(* IEC 61131-3 sources: plc-iiot-stack/tests/POUs/F_TestContains, 2 files *)

(* ---- F_TestContains.decl.st ---- *)
// Назначение: для тестов — содержит ли текст длиной до MQTT_PAYLOAD_LEN подстроку sPart (стандартная
//             FIND работает только со строками до 255 символов).
// Автор:      kr0nsch
// Версия:     0.1.0
// Документ:   docs/TEST_REPORT.md
FUNCTION F_TestContains : BOOL
VAR_IN_OUT CONSTANT
    // lint:allow STL007 параметр VAR_IN_OUT CONSTANT — ссылка только для чтения, а не константа
    sText : STRING(GVL_Const.MQTT_PAYLOAD_LEN);
END_VAR
VAR_INPUT
    sPart : STRING(255);
END_VAR
VAR
    uiTextLen : UINT;
    uiPartLen : UINT;
    uiStart : UINT;
    uiIdx : UINT;
    xMatch : BOOL;
END_VAR

(* ---- F_TestContains.impl.st ---- *)
uiPartLen := INT_TO_UINT(LEN(sPart));
uiTextLen := 0;
WHILE uiTextLen < GVL_Const.MQTT_PAYLOAD_LEN AND_THEN sText[uiTextLen] <> 0 DO
    uiTextLen := uiTextLen + 1;
END_WHILE
IF uiPartLen = 0 THEN
    F_TestContains := TRUE;
    RETURN;
END_IF
IF uiPartLen > uiTextLen THEN
    RETURN;
END_IF
FOR uiStart := 0 TO uiTextLen - uiPartLen DO
    xMatch := TRUE;
    FOR uiIdx := 0 TO uiPartLen - 1 DO
        IF sText[uiStart + uiIdx] <> sPart[uiIdx] THEN
            xMatch := FALSE;
            EXIT;
        END_IF
    END_FOR
    IF xMatch THEN
        F_TestContains := TRUE;
        RETURN;
    END_IF
END_FOR
